{attribute 'qualified_only'}
{attribute 'strict'}
TYPE WheelSide :
(
	LEFT := 0,
	RIGHT
);
END_TYPE

(* stored: Version 1.1.0.1, ProductVersion 3.1.4026.12
   DUT WheelSide: Id {df027a90-f2d2-5faf-85eb-7778b97dc1da} *)
